DATA_BLOCK "FRK_ModelStore"
{ S7_Optimized_Access := 'TRUE' }
VERSION : 0.1
NON_RETAIN
VAR RETAIN
    Rows {ExternalAccessible := 'False'; ExternalVisible := 'False'; ExternalWritable := 'False'} : Array[1..1] of "FRK_ModelCatalog";
END_VAR
BEGIN
END_DATA_BLOCK
